// TIA Portal V20 export
DATA_BLOCK "DB_data_ctena"   // DB7
{ S7_Optimized_Access := 'TRUE' }
// stored: MemoryReserve 100
   VAR
      array_of_byte : Array[0..150] of Byte;
      array_of_char : Array[0..150] of Char;
      cteny_string : String[150];
      upraveny : String[150];
   END_VAR
BEGIN
END_DATA_BLOCK
